Fanuc KAREL source: kt00052.KL

-- PROVISIONAL review KL for V1013-1; original PC SHA256 53dd9d7ab0255920faf4693110ac9b96ed305547adc8a2364c07221df09d6c28
-- Incomplete behavior may be omitted. Consult companion uncertainty JSON. Do not deploy.
PROGRAM KT00052
%NOLOCKGROUP
VAR
  R2 : REAL
  OUT : REAL
-- UNRESOLVED_DECL Y1 type=002018
BEGIN
  -- UNRESOLVED_PC offsets 5-19; opcodes 2E,22,9D,33,B2
  -- UNRESOLVED_PC offsets 24-35; opcodes 2E,23
  -- UNRESOLVED_PC offsets 40-65; opcodes 22,9D,33,B1,21,29,64,29,6A,23
  -- UNRESOLVED_PC offsets 70-74; opcodes 7F
END KT00052
